// TIA Portal V21 export
// export: Created 2000-01-01T00:00:00.0000000Z, ExportSetting None
TYPE "UDT_HMI_ModbusPoller"
   STRUCT
      bEnablePoll { ExternalWritable := 'False'} : Bool;   // HMI轮询总使能开关
      bResetStats { ExternalWritable := 'False'} : Bool;   // HMI清零通信统计与故障计数
      iMaxStationCount { ExternalWritable := 'False'} : Int;   // 参与轮询的从站总数 (1..8，默认 4)
      iMaxRetryCount { ExternalWritable := 'False'} : Int;   // 单站超时最大重试次数 (0..5，默认 3)
      tReplyTimeout { ExternalWritable := 'False'} : Time;   // 单次请求响应超时时间（默认 T#1s）
      tInterFrameDelay { ExternalWritable := 'False'} : Time;   // 帧间静默轮询间隔时间（默认 T#50ms）
      iActiveStationIdx { ExternalWritable := 'False'} : Int;   // 状态反馈：当前正在轮询的站索引 (1..8)
      diSuccessCount { ExternalWritable := 'False'} : DInt;   // 状态反馈：累计成功通信次数
      diErrorCount { ExternalWritable := 'False'} : DInt;   // 状态反馈：累计失败通信次数
      bAnyStationFault { ExternalWritable := 'False'} : Bool;   // 状态反馈：存在从站掉线报警
      wStatus { ExternalWritable := 'False'} : Word;   // 状态码：16#0000一轮完成, 16#7000未激活, 16#7002轮询中, 16#8401从站超时掉线
   END_STRUCT;
END_TYPE
